// TIA Portal V19 export
// export: Created 2026-10-15T09:44:24.3054294Z, ExportSetting WithDefaults, DisplayName Totally Integrated Automation Portal, DisplayVersion V19, DisplayName TIA Portal Openness, DisplayVersion V19, DisplayName TIA Portal Version Control Interface, DisplayVersion V19, DisplayName STEP 7 Professional, DisplayVersion V19, DisplayName STEP 7 Safety, DisplayVersion V19, DisplayName WinCC Basic/Comfort/Advanced, DisplayVersion V19, DisplayName WinCC Unified, DisplayVersion V19
FUNCTION "ROLL_PB15" : Void   // FC23, SCL
{ S7_Optimized_Access := 'TRUE' }
VERSION : 0.1
// stored: AutoNumber true, IsIECCheckEnabled false, SetENOAutomatically false, UDAEnableTagReadback false
   VAR_TEMP
      r : Bool;
      a1 : Word;
      a2 : Word;
      activeDataBlock : Int;
      comparisonResults : Array[0..0] of Bool;
   END_VAR
BEGIN

   #r := FALSE;
   #a1 := W#16#0000;
   #a2 := W#16#0000;
   #activeDataBlock := 0;
   // PB15, STEP 5 network 1
   #r := ((NOT "ROLL_IO".Output[113, 2]) AND "ROLL_IO".Output[113, 3] AND "ROLL_IO".Input[123, 4]);
   IF #r THEN
       "ROLL_State".M[70, 2] := TRUE;
   END_IF;
   #r := (((NOT "ROLL_IO".Input[123, 4]) AND "ROLL_IO".Input[123, 5]) OR "ROLL_State".M[73, 7]);
   IF #r THEN
       "ROLL_State".M[70, 2] := FALSE;
   END_IF;
   // PB15, STEP 5 network 2
   #r := ((((NOT "ROLL_State".M[20, 2]) AND "ROLL_IO".Input[123, 6] AND "ROLL_State".M[74, 0]) OR "ROLL_State".M[71, 0]) AND "ROLL_IO".Output[113, 2] AND "ROLL_IO".Input[124, 1] AND "ROLL_IO".Input[124, 4]);
   IF #r THEN
       "ROLL_State".M[70, 3] := TRUE;
   END_IF;
   #r := (((NOT "ROLL_IO".Input[123, 5]) AND (NOT "ROLL_IO".Input[123, 6])) OR "ROLL_State".M[73, 7]);
   IF #r THEN
       "ROLL_State".M[70, 3] := FALSE;
   END_IF;
   // PB15, STEP 5 network 3
   #r := ((NOT "ROLL_State".M[16, 0]) AND (NOT "ROLL_State".M[16, 1]) AND (NOT "ROLL_State".M[16, 4]) AND (NOT "ROLL_State".M[71, 1]) AND "ROLL_IO".Input[123, 1] AND "ROLL_State".M[191, 4] AND "ROLL_State".M[31, 4] AND "ROLL_State".S5Timers[45].Q);
   IF #r THEN
       "ROLL_State".M[70, 4] := TRUE;
   END_IF;
   #r := ((NOT "ROLL_IO".Input[123, 1]) OR "ROLL_State".M[73, 7]);
   IF #r THEN
       "ROLL_State".M[70, 4] := FALSE;
   END_IF;
   // PB15, STEP 5 network 4
   #r := "ROLL_IO".Input[123, 6];
   IF #r THEN
       "ROLL_State".M[70, 5] := TRUE;
   END_IF;
   #r := ("ROLL_IO".Input[125, 0] OR "ROLL_State".M[73, 7]);
   IF #r THEN
       "ROLL_State".M[70, 5] := FALSE;
   END_IF;
   // PB15, STEP 5 network 5
   #r := ((NOT "ROLL_IO".Input[125, 1]) AND "ROLL_IO".Output[113, 4] AND "ROLL_IO".Input[125, 0]);
   IF #r THEN
       "ROLL_State".M[70, 6] := TRUE;
   END_IF;
   #r := (("ROLL_IO".Output[113, 5] AND "ROLL_IO".Input[125, 1]) OR "ROLL_State".M[73, 7]);
   IF #r THEN
       "ROLL_State".M[70, 6] := FALSE;
   END_IF;
   // PB15, STEP 5 network 6
   #r := ((NOT "ROLL_State".M[71, 1]) AND "ROLL_IO".Input[123, 1] AND "ROLL_State".S5Timers[45].Q);
   IF #r THEN
       "ROLL_State".M[70, 7] := TRUE;
   END_IF;
   #r := ("ROLL_IO".Input[123, 4] OR "ROLL_State".M[73, 7]);
   IF #r THEN
       "ROLL_State".M[70, 7] := FALSE;
   END_IF;
   // PB15, STEP 5 network 7
   #r := ("ROLL_IO".Output[113, 3] AND "ROLL_IO".Input[123, 5]);
   IF #r THEN
       "ROLL_State".M[71, 0] := TRUE;
   END_IF;
   #r := ("ROLL_State".M[70, 3] OR "ROLL_State".M[73, 7]);
   IF #r THEN
       "ROLL_State".M[71, 0] := FALSE;
   END_IF;
   // PB15, STEP 5 network 8
   #r := ((NOT "ROLL_State".M[190, 6]) AND (NOT "ROLL_State".M[28, 4]) AND ("ROLL_State".M[20, 1] OR "ROLL_State".M[20, 2]) AND "ROLL_IO".Input[0, 1] AND "ROLL_State".M[190, 5]);
   "ROLL_State".M[74, 0] := #r;
   // PB15, STEP 5 network 9
   RETURN;
END_FUNCTION
